        bool bMarked
        jointRx jJointRx = {j1=-132.269491, j2=127.123938, j3=-106.855674, j4=181.429188, j5=21.342688, j6=130.953129}
        pointRx pInter
        paraItem pParaItem
          [0]
            bool bSafePoint
            ifItem iIfItem
              [0]
                bool bANDOR[2]
                num nSigIndex[3]
                num nSigType[3]
                num nValue[3]
            mdesc mMdesc
            num nActionIndex = 42
            num nDelay
            num nMoveType = 1
            num nPercentage
            num nSigValue = 1
        pointRx pPointRx[2] = {x=-320.674662, y=-420.382638, z=642.0718966, rx=-1.140431, ry=0.333681, rz=-179.976981, shoulder=lefty, elbow=enegative, wrist=wpositive}
        string sID
      [45]
        bool bMarked
        jointRx jJointRx = {j1=-142.441106, j2=120.824327, j3=-88.705493, j4=181.282913, j5=33.0850501, j6=141.380041}
        pointRx pInter
        paraItem pParaItem
          [0]
            bool bSafePoint
            ifItem iIfItem
              [0]
                bool bANDOR[2]
                num nSigIndex[3]
                num nSigType[3]
                num nValue[3]
            mdesc mMdesc
            num nActionIndex = 42
            num nDelay
            num nMoveType = 1
            num nPercentage
            num nSigValue = 1
        pointRx pPointRx[2] = {x=-474.689621, y=-420.382631, z=642.0718894, rx=-1.140119, ry=0.333784, rz=-179.976923, shoulder=lefty, elbow=enegative, wrist=wpositive}
        string sID
      [46]
        bool bMarked
        jointRx jJointRx = {j1=-138.108258, j2=121.207146, j3=-89.710766, j4=181.162609, j5=32.51161, j6=137.142341}
        pointRx pInter
        paraItem pParaItem
          [0]
            bool bSafePoint
            ifItem iIfItem
              [0]
                bool bANDOR[2]
                num nSigIndex[3]
                num nSigType[3]
                num nValue[3]
            mdesc mMdesc
            num nActionIndex = 42
            num nDelay
            num nMoveType = 1
            num nPercentage
            num nSigValue = 1
        pointRx pPointRx[2] = {x=-436.796862, y=-451.644484, z=642.07189, rx=-1.139469, ry=0.334472, rz=-179.976638, shoulder=lefty, elbow=enegative, wrist=wpositive}
        string sID
      [47]
        bool bMarked
        jointRx jJointRx = {j1=-127.70596, j2=126.693595, j3=-105.454305, j4=181.135682, j5=22.350888, j6=126.671469}
        pointRx pInter
        paraItem pParaItem
          [0]
            bool bSafePoint
            ifItem iIfItem
              [0]
                bool bANDOR[2]
                num nSigIndex[3]
                num nSigType[3]
                num nValue[3]
            mdesc mMdesc
            num nActionIndex = 42
            num nDelay
            num nMoveType = 1
            num nPercentage
            num nSigValue = 1
        pointRx pPointRx[2] = {x=-290.683508, y=-451.609469, z=642.07191, rx=-1.140457, ry=0.335724, rz=-179.976594, shoulder=lefty, elbow=enegative, wrist=wpositive}
        string sID
      [48]
        bool bMarked
        jointRx jJointRx = {j1=-77.238254, j2=129.340507, j3=-114.913945, j4=177.831104, j5=15.475362, j6=79.35375}
        pointRx pInter
        paraItem pParaItem
          [0]
            bool bSafePoint
            ifItem iIfItem
              [0]
                bool bANDOR[2]
                num nSigIndex[3]
                num nSigType[3]
                num nValue[3]
            mdesc mMdesc
            num nActionIndex = 42
            num nDelay
            num nMoveType = 1
            num nPercentage
            num nSigValue = 1
        pointRx pPointRx[2] = {x=158.729452, y=-451.609464, z=642.0719065, rx=-1.140389, ry=0.334964, rz=-179.976748, shoulder=lefty, elbow=enegative, wrist=wpositive}
        string sID
      [49]
        bool bMarked
        jointRx jJointRx = {j1=-63.488687, j2=124.208026, j3=-97.940675, j4=178.228458, j5=27.14867, j6=65.0910716}
        pointRx pInter
        paraItem pParaItem
          [0]
            bool bSafePoint
            ifItem iIfItem
              [0]
                bool bANDOR[2]
                num nSigIndex[3]
                num nSigType[3]
                num nValue[3]
            mdesc mMdesc
            num nActionIndex = 42
            num nDelay
            num nMoveType = 1
            num nPercentage
            num nSigValue = 1
        pointRx pPointRx[2] = {x=310.830797, y=-495.30753, z=642.0718875, rx=-1.139453, ry=0.33486, rz=-179.976891, shoulder=lefty, elbow=enegative, wrist=wpositive}
        string sID
      [50]
        bool bMarked
        jointRx jJointRx = {j1=-78.0579912, j2=127.559769, j3=-108.316642, j4=178.378161, j5=20.297351, j6=79.604006}
        pointRx pInter
        paraItem pParaItem
          [0]
            bool bSafePoint
            ifItem iIfItem
              [0]
                bool bANDOR[2]
                num nSigIndex[3]
                num nSigType[3]
                num nValue[3]
            mdesc mMdesc
            num nActionIndex = 42
            num nDelay
            num nMoveType = 1
            num nPercentage
            num nSigValue = 1
        pointRx pPointRx[2] = {x=160.873249, y=-495.272541, z=642.0719096, rx=-1.140489, ry=0.333782, rz=-179.976981, shoulder=lefty, elbow=enegative, wrist=wpositive}
        string sID
      [51]
        bool bMarked
        jointRx jJointRx = {j1=-83.970136, j2=129.00855342, j3=-113.590578, j4=181.751291, j5=14.32041, j6=-96.622719}
        pointRx pInter
        paraItem pParaItem
          [0]
            bool bSafePoint
            ifItem iIfItem
              [0]
                bool bANDOR[2]
                num nSigIndex[3]
                num nSigType[3]
                num nValue[3]
            mdesc mMdesc
            num nActionIndex = 42
            num nDelay
            num nMoveType = 1
            num nPercentage
            num nSigValue = 1
        pointRx pPointRx[2] = {x=98.789636, y=-495.232609, z=642.0875542, rx=1.143362, ry=-0.31475, rz=1.103019, shoulder=lefty, elbow=enegative, wrist=wpositive}
        string sID
      [52]
        bool bMarked
        jointRx jJointRx = {j1=-101.251443, j2=129.329307, j3=-114.876217, j4=180.377122, j5=13.270505, j6=-78.0149862}
        pointRx pInter
        paraItem pParaItem
          [0]
            bool bSafePoint
            ifItem iIfItem
              [0]
                bool bANDOR[2]
                num nSigIndex[3]
                num nSigType[3]
                num nValue[3]
            mdesc mMdesc
            num nActionIndex = 42
            num nDelay
            num nMoveType = 1
            num nPercentage
            num nSigValue = 1
        pointRx pPointRx[2] = {x=-48.311282, y=-495.232554, z=642.0875543, rx=1.143247, ry=-0.315683, rz=1.102879, shoulder=lefty, elbow=enegative, wrist=wpositive}
        string sID
      [53]
        bool bMarked
        jointRx jJointRx = {j1=-117.974593, j2=127.746571, j3=-108.963712, j4=179.150072, j5=17.626951, j6=-60.118292}
        pointRx pInter
        paraItem pParaItem
          [0]
            bool bSafePoint
            ifItem iIfItem
              [0]
                bool bANDOR[2]
                num nSigIndex[3]
                num nSigType[3]
                num nValue[3]
            mdesc mMdesc
            num nActionIndex = 42
            num nDelay
            num nMoveType = 1
            num nPercentage
            num nSigValue = 1
        pointRx pPointRx[2] = {x=-203.879984, y=-495.232578, z=642.0875477, rx=1.143192, ry=-0.315734, rz=1.102838, shoulder=lefty, elbow=enegative, wrist=wpositive}
        string sID
      [54]
        bool bMarked
        jointRx jJointRx = {j1=-130.30363, j2=123.943868, j3=-97.190977, j4=178.849142, j5=25.681002, j6=-47.564193}
        pointRx pInter
        paraItem pParaItem
          [0]
            bool bSafePoint
            ifItem iIfItem
              [0]
                bool bANDOR[2]
                num nSigIndex[3]
                num nSigType[3]
                num nValue[3]
            mdesc mMdesc
            num nActionIndex = 42
            num nDelay
            num nMoveType = 1
            num nPercentage
            num nSigValue = 1
        pointRx pPointRx[2] = {x=-348.772288, y=-495.232559, z=642.0875407, rx=1.143488, ry=-0.315869, rz=1.102811, shoulder=lefty, elbow=enegative, wrist=wpositive}
        string sID
      [55]
        bool bMarked
        jointRx jJointRx = {j1=-87.553471, j2=145.12737, j3=-83.0900686, j4=182.117938, j5=63.691767, j6=-64.957345}
        pointRx pInter
        paraItem pParaItem
          [0]
            bool bSafePoint
            ifItem iIfItem
              [0]
                bool bANDOR[2]
                num nSigIndex[3]
                num nSigType[3]
                num nValue[3]
            mdesc mMdesc
            num nActionIndex = 42
            num nDelay
            num nMoveType = 1
            num nPercentage
            num nSigValue = 1
        pointRx pPointRx[2] = {x=61.326125, y=-652.062172, z=350.121525, rx=-1.556374, ry=-1.966704, rz=28.428639, shoulder=lefty, elbow=enegative, wrist=wpositive}
        string sID
    string sID
  [Position8_point_blow]
    num nFrameIndex
    num nMoveID
    num nToolIndex
    pointItem pPointItem[50]
      [0]
        bool bMarked
        jointRx jJointRx
        pointRx pInter
        paraItem pParaItem
          [0]
            bool bSafePoint
            ifItem iIfItem
              [0]
                bool bANDOR[2]
                num nSigIndex[3]
                num nSigType[3]
                num nValue[3]
            mdesc mMdesc
            num nActionIndex = 43
            num nDelay
            num nMoveType = 4
            num nPercentage
            num nSigValue = 1
        pointRx pPointRx[2]
        string sID
      [1]
        bool bMarked
        jointRx jJointRx = {j1=-87.553471, j2=145.12737, j3=-83.0900679, j4=182.117938, j5=63.691768, j6=-64.957345}
        pointRx pInter
        paraItem pParaItem
          [0]
            bool bSafePoint
            ifItem iIfItem
              [0]
                bool bANDOR[2]
                num nSigIndex[3]
                num nSigType[3]
                num nValue[3]
            mdesc mMdesc
            num nActionIndex = 42
            num nDelay
            num nMoveType = 1
            num nPercentage
            num nSigValue = 1
        pointRx pPointRx[2] = {x=61.326125, y=-652.062172, z=350.121525, rx=-1.556374, ry=-1.966704, rz=28.428639, shoulder=lefty, elbow=enegative, wrist=wpositive}
        string sID
      [2]
        bool bMarked
        jointRx jJointRx = {j1=-58.11069, j2=109.524278, j3=-71.857715, j4=179.347561, j5=40.141515, j6=-122.34843}
        pointRx pInter
        paraItem pParaItem
          [0]
            bool bSafePoint
            ifItem iIfItem
              [0]
                bool bANDOR[2]
                num nSigIndex[3]
                num nSigType[3]
                num nValue[3]
            mdesc mMdesc
            num nActionIndex = 42
            num nDelay
            num nMoveType = 1
            num nPercentage
            num nSigValue = 1
        pointRx pPointRx[2] = {x=409.39132, y=-556.393527, z=693.904783, rx=-2.322296, ry=-0.948981, rz=-0.986203, shoulder=lefty, elbow=enegative, wrist=wpositive}
        string sID
      [3]
        bool bMarked
        jointRx jJointRx = {j1=-66.225547, j2=113.999088, j3=-83.778734, j4=179.876465, j5=32.728091, j6=-114.636276}
        pointRx pInter
        paraItem pParaItem
          [0]
            bool bSafePoint
            ifItem iIfItem
              [0]
                bool bANDOR[2]
                num nSigIndex[3]
                num nSigType[3]
                num nValue[3]
            mdesc mMdesc
            num nActionIndex = 42
            num nDelay
            num nMoveType = 1
            num nPercentage
            num nSigValue = 1
        pointRx pPointRx[2] = {x=300.386557, y=-556.417777, z=693.904772, rx=-2.32202, ry=-0.949536, rz=-0.986453, shoulder=lefty, elbow=enegative, wrist=wpositive}
        string sID
      [4]
        bool bMarked
        jointRx jJointRx = {j1=-76.687433, j2=116.715992, j3=-91.802088, j4=180.847193, j5=27.394171, j6=-105.0405035}
        pointRx pInter
        paraItem pParaItem
          [0]
            bool bSafePoint
            ifItem iIfItem
              [0]
                bool bANDOR[2]
                num nSigIndex[3]
                num nSigType[3]
                num nValue[3]
            mdesc mMdesc
            num nActionIndex = 42
            num nDelay
            num nMoveType = 1
            num nPercentage
            num nSigValue = 1
        pointRx pPointRx[2] = {x=180.521932, y=-560.5436, z=693.904726, rx=-2.321521, ry=-0.949691, rz=-0.986547, shoulder=lefty, elbow=enegative, wrist=wpositive}
        string sID
      [5]
        bool bMarked
        jointRx jJointRx = {j1=-85.620281, j2=117.92465, j3=-95.696322, j4=181.846877, j5=24.627005, j6=-97.0419871}
        pointRx pInter
        paraItem pParaItem
          [0]
            bool bSafePoint
            ifItem iIfItem
              [0]
                bool bANDOR[2]
                num nSigIndex[3]
                num nSigType[3]
                num nValue[3]
            mdesc mMdesc
            num nActionIndex = 42
            num nDelay
            num nMoveType = 1
            num nPercentage
            num nSigValue = 1
        pointRx pPointRx[2] = {x=86.341042, y=-560.508796, z=693.904766, rx=-2.321719, ry=-0.949521, rz=-0.986489, shoulder=lefty, elbow=enegative, wrist=wpositive}
        string sID
      [6]
        bool bMarked
        jointRx jJointRx = {j1=-101.0757166, j2=116.15458, j3=-90.0727261, j4=182.913944, j5=28.207981, j6=-82.484873}
        pointRx pInter
        paraItem pParaItem
          [0]
            bool bSafePoint
            ifItem iIfItem
              [0]
                bool bANDOR[2]
                num nSigIndex[3]
                num nSigType[3]
                num nValue[3]
            mdesc mMdesc
            num nActionIndex = 42
            num nDelay
            num nMoveType = 1
            num nPercentage
            num nSigValue = 1
        pointRx pPointRx[2] = {x=-77.997367, y=-596.182081, z=693.904723, rx=-2.320616, ry=-0.948845, rz=-0.986256, shoulder=lefty, elbow=enegative, wrist=wpositive}
        string sID
      [7]
        bool bMarked
        jointRx jJointRx = {j1=-100.388707, j2=113.501769, j3=-82.38876, j4=182.465739, j5=33.248966, j6=-82.665703}
        pointRx pInter
        paraItem pParaItem
          [0]
            bool bSafePoint
            ifItem iIfItem
              [0]
                bool bANDOR[2]
                num nSigIndex[3]
                num nSigType[3]
                num nValue[3]
            mdesc mMdesc
            num nActionIndex = 42
            num nDelay
            num nMoveType = 1
            num nPercentage
            num nSigValue = 1
        pointRx pPointRx[2] = {x=-77.997368, y=-637.319122, z=693.904719, rx=-2.320623, ry=-0.948795, rz=-0.986246, shoulder=lefty, elbow=enegative, wrist=wpositive}
        string sID
      [8]
        bool bMarked
        jointRx jJointRx = {j1=-112.569059, j2=111.105712, j3=-75.937343, j4=182.939146, j5=36.983748, j6=-70.774258}
        pointRx pInter
        paraItem pParaItem
          [0]
            bool bSafePoint
            ifItem iIfItem
              [0]
                bool bANDOR[2]
                num nSigIndex[3]
                num nSigType[3]
                num nValue[3]
            mdesc mMdesc
            num nActionIndex = 42
            num nDelay
            num nMoveType = 1
            num nPercentage
            num nSigValue = 1
        pointRx pPointRx[2] = {x=-227.428005, y=-637.284544, z=693.904751, rx=-2.321115, ry=-0.949679, rz=-0.986554, shoulder=lefty, elbow=enegative, wrist=wpositive}
        string sID
      [9]
        bool bMarked
        jointRx jJointRx = {j1=-113.957376, j2=114.00103433, j3=-83.784205, j4=183.416468, j5=32.000017554, j6=-69.935449}
        pointRx pInter
        paraItem pParaItem
          [0]
            bool bSafePoint
            ifItem iIfItem
              [0]
                bool bANDOR[2]
                num nSigIndex[3]
                num nSigType[3]
                num nValue[3]
            mdesc mMdesc
            num nActionIndex = 42
            num nDelay
            num nMoveType = 1
            num nPercentage
            num nSigValue = 1
        pointRx pPointRx[2] = {x=-227.392618, y=-596.00613787, z=693.904773, rx=-2.322353, ry=-0.948517, rz=-0.986316, shoulder=lefty, elbow=enegative, wrist=wpositive}
        string sID
      [10]
        bool bMarked
        jointRx jJointRx = {j1=-131.107782, j2=122.205733, j3=-114.25278, j4=193.937243, j5=9.352415, j6=-63.640524}
        pointRx pInter
        paraItem pParaItem
          [0]
            bool bSafePoint
            ifItem iIfItem
              [0]
                bool bANDOR[2]
                num nSigIndex[3]
                num nSigType[3]
                num nValue[3]
            mdesc mMdesc
            num nActionIndex = 42
            num nDelay
            num nMoveType = 1
            num nPercentage
            num nSigValue = 1
        pointRx pPointRx[2] = {x=-278.571769, y=-365.527339, z=693.923849, rx=-2.325235, ry=-0.948268, rz=-0.986383, shoulder=lefty, elbow=enegative, wrist=wpositive}
        string sID
      [11]
        bool bMarked
        jointRx jJointRx = {j1=-135.395911, j2=104.707172, j3=-76.504799, j4=184.753699, j5=29.243911, j6=-49.740588}
        pointRx pInter
        paraItem pParaItem
          [0]
            bool bSafePoint
            ifItem iIfItem
              [0]
                bool bANDOR[2]
                num nSigIndex[3]
                num nSigType[3]
                num nValue[3]
            mdesc mMdesc
            num nActionIndex = 42
            num nDelay
            num nMoveType = 1
            num nPercentage
            num nSigValue = 1
        pointRx pPointRx[2] = {x=-444.435288, y=-480.130514, z=766.167371, rx=-2.324241, ry=-0.947818, rz=-0.986236, shoulder=lefty, elbow=enegative, wrist=wpositive}
        string sID
      [12]
        bool bMarked
        jointRx jJointRx = {j1=-134.796217, j2=92.950158, j3=-65.644872, j4=184.86577, j5=28.374058, j6=-50.474125}
        pointRx pInter
        paraItem pParaItem
          [0]
            bool bSafePoint
            ifItem iIfItem
              [0]
                bool bANDOR[2]
                num nSigIndex[3]
                num nSigType[3]
                num nValue[3]
            mdesc mMdesc
            num nActionIndex = 42
            num nDelay
            num nMoveType = 1
            num nPercentage
            num nSigValue = 1
        pointRx pPointRx[2] = {x=-444.435359, y=-489.966612, z=855.290958, rx=-2.324744, ry=-0.947384, rz=-0.986218, shoulder=lefty, elbow=enegative, wrist=wpositive}
        string sID
      [13]
        bool bMarked
        jointRx jJointRx = {j1=-136.173853, j2=87.871737, j3=-63.130701, j4=185.374273, j5=25.767564, j6=-49.65473}
        pointRx pInter
        paraItem pParaItem
          [0]
            bool bSafePoint
            ifItem iIfItem
              [0]
                bool bANDOR[2]
                num nSigIndex[3]
                num nSigType[3]
                num nValue[3]
            mdesc mMdesc
            num nActionIndex = 42
            num nDelay
            num nMoveType = 1
            num nPercentage
            num nSigValue = 1
        pointRx pPointRx[2] = {x=-444.435358, y=-467.674325, z=901.291627, rx=-2.325949, ry=-0.946701, rz=-0.986341, shoulder=lefty, elbow=enegative, wrist=wpositive}
        string sID
      [14]
        bool bMarked
        jointRx jJointRx = {j1=-141.164951, j2=86.59666, j3=-69.357957, j4=187.756915, j5=18.114888, j6=-47.194082}
        pointRx pInter
        paraItem pParaItem
          [0]
            bool bSafePoint
            ifItem iIfItem
              [0]
                bool bANDOR[2]
                num nSigIndex[3]
                num nSigType[3]
                num nValue[3]
            mdesc mMdesc
            num nActionIndex = 42
            num nDelay
            num nMoveType = 1
            num nPercentage
            num nSigValue = 1
        pointRx pPointRx[2] = {x=-444.435342, y=-395.0345733, z=930.658223, rx=-2.325698, ry=-0.946616, rz=-0.986323, shoulder=lefty, elbow=enegative, wrist=wpositive}
        string sID
      [15]
        bool bMarked
        jointRx jJointRx = {j1=-150.996048, j2=88.749744, j3=-81.786263, j4=199.00922873, j5=7.675391, j6=-48.828489}
        pointRx pInter
        paraItem pParaItem
          [0]
            bool bSafePoint
            ifItem iIfItem
              [0]
                bool bANDOR[2]
                num nSigIndex[3]
                num nSigType[3]
                num nValue[3]
            mdesc mMdesc
            num nActionIndex = 42
            num nDelay
            num nMoveType = 1
            num nPercentage
            num nSigValue = 1
        pointRx pPointRx[2] = {x=-444.435068, y=-278.693508, z=930.65815, rx=-2.325239, ry=-0.948289, rz=-0.986304, shoulder=lefty, elbow=enegative, wrist=wpositive}
        string sID
      [16]
        bool bMarked
        jointRx jJointRx = {j1=-136.944318, j2=108.102124, j3=-81.594441, j4=185.0858237, j5=27.496189, j6=-48.554881}
        pointRx pInter
        paraItem pParaItem
          [0]
            bool bSafePoint
            ifItem iIfItem
              [0]
                bool bANDOR[2]
                num nSigIndex[3]
                num nSigType[3]
                num nValue[3]
            mdesc mMdesc
            num nActionIndex = 42
            num nDelay
            num nMoveType = 1
            num nPercentage
            num nSigValue = 1
        pointRx pPointRx[2] = {x=-444.435337, y=-455.673073, z=747.789181, rx=-2.325621, ry=-0.946829, rz=-0.986212, shoulder=lefty, elbow=enegative, wrist=wpositive}
        string sID
      [17]
        bool bMarked
        jointRx jJointRx = {j1=-133.102266, j2=114.394979, j3=-110.124586, j4=185.156231, j5=6.735085, j6=-104.330607}
        pointRx pInter
        paraItem pParaItem
          [0]
            bool bSafePoint
            ifItem iIfItem
              [0]
                bool bANDOR[2]
                num nSigIndex[3]
                num nSigType[3]
                num nValue[3]
            mdesc mMdesc
            num nActionIndex = 42
            num nDelay
            num nMoveType = 1
            num nPercentage
            num nSigValue = 1
        pointRx pPointRx[2] = {x=-273.0764108, y=-357.254112, z=747.804416, rx=-2.192889, ry=1.224247, rz=-52.275755, shoulder=lefty, elbow=enegative, wrist=wpositive}
        string sID
      [18]
        bool bMarked
        jointRx jJointRx = {j1=-117.270513, j2=113.78497, j3=-104.717978, j4=179.481532, j5=11.577034, j6=-114.962229}
        pointRx pInter
        paraItem pParaItem
          [0]
            bool bSafePoint
            ifItem iIfItem
              [0]
                bool bANDOR[2]
                num nSigIndex[3]
                num nSigType[3]
                num nValue[3]
            mdesc mMdesc
            num nActionIndex = 42
            num nDelay
            num nMoveType = 1
            num nPercentage
            num nSigValue = 1
        pointRx pPointRx[2] = {x=-176.508441, y=-453.51729, z=747.804419, rx=-2.183299, ry=1.242081, rz=-52.719273, shoulder=lefty, elbow=enegative, wrist=wpositive}
        string sID
      [19]
        bool bMarked
        jointRx jJointRx = {j1=-109.137554, j2=109.619736, j3=-86.542307, j4=178.941557, j5=25.551631, j6=-122.640865}
        pointRx pInter
        paraItem pParaItem
          [0]
            bool bSafePoint
            ifItem iIfItem
              [0]
                bool bANDOR[2]
                num nSigIndex[3]
                num nSigType[3]
                num nValue[3]
            mdesc mMdesc
            num nActionIndex = 42
            num nDelay
            num nMoveType = 1
            num nPercentage
            num nSigValue = 1
        pointRx pPointRx[2] = {x=-144.182021, y=-580.158289, z=747.804426, rx=-2.184454, ry=1.240986, rz=-52.719545, shoulder=lefty, elbow=enegative, wrist=wpositive}
        string sID
      [20]
        bool bMarked
        jointRx jJointRx = {j1=-105.96936, j2=113.946894, j3=-105.873919, j4=176.762051, j5=10.531462, j6=-123.577788}
        pointRx pInter
        paraItem pParaItem
          [0]
            bool bSafePoint
            ifItem iIfItem
              [0]
                bool bANDOR[2]
                num nSigIndex[3]
                num nSigType[3]
                num nValue[3]
            mdesc mMdesc
            num nActionIndex = 42
            num nDelay
            num nMoveType = 1
            num nPercentage
            num nSigValue = 1
        pointRx pPointRx[2] = {x=-78.145175, y=-473.574291, z=747.804414, rx=-2.185277, ry=1.240398, rz=-52.719616, shoulder=lefty, elbow=enegative, wrist=wpositive}
        string sID
      [21]
        bool bMarked
        jointRx jJointRx = {j1=-100.135452, j2=114.341428, j3=-109.460145, j4=173.401757, j5=7.298155, j6=-126.0452472}
        pointRx pInter
        paraItem pParaItem
          [0]
            bool bSafePoint
            ifItem iIfItem
              [0]
                bool bANDOR[2]
                num nSigIndex[3]
                num nSigType[3]
                num nValue[3]
            mdesc mMdesc
            num nActionIndex = 42
            num nDelay
            num nMoveType = 1
            num nPercentage
            num nSigValue = 1
        pointRx pPointRx[2] = {x=-23.263146, y=-455.736187, z=747.804388, rx=-2.18503, ry=1.240118, rz=-52.719596, shoulder=lefty, elbow=enegative, wrist=wpositive}
        string sID
      [22]
        bool bMarked
        jointRx jJointRx = {j1=-100.135452, j2=114.341428, j3=-109.460145, j4=173.401757, j5=7.298155, j6=-126.0452472}
        pointRx pInter
        paraItem pParaItem
          [0]
            bool bSafePoint
            ifItem iIfItem
              [0]
                bool bANDOR[2]
                num nSigIndex[3]
                num nSigType[3]
                num nValue[3]
            mdesc mMdesc
            num nActionIndex = 42
            num nDelay
            num nMoveType
            num nPercentage
            num nSigValue = 1
        pointRx pPointRx[2] = {x=-23.263146, y=-455.736187, z=747.804388, rx=-2.18503, ry=1.240118, rz=-52.719596, shoulder=lefty, elbow=enegative, wrist=wpositive}
        string sID
      [23]
        bool bMarked
        jointRx jJointRx = {j1=-106.631553, j2=109.786963, j3=-134.970625, j4=184.819916, j5=-24.691551, j6=-80.199638}
        pointRx pInter
        paraItem pParaItem
          [0]
            bool bSafePoint
            ifItem iIfItem
              [0]
                bool bANDOR[2]
                num nSigIndex[3]
                num nSigType[3]
                num nValue[3]
            mdesc mMdesc
            num nActionIndex = 42
            num nDelay
            num nMoveType
            num nPercentage
            num nSigValue = 1
        pointRx pPointRx[2] = {x=-10.865105, y=-272.383063, z=740.397718, rx=0.0307126, ry=2.090166, rz=-2.46071, shoulder=lefty, elbow=enegative, wrist=wnegative}
        string sID
      [24]
        bool bMarked
        jointRx jJointRx = {j1=-81.325877, j2=110.844378, j3=-133.586221, j4=185.246198, j5=-23.174992, j6=-105.96506}
        pointRx pInter
        paraItem pParaItem
          [0]
            bool bSafePoint
            ifItem iIfItem
              [0]
                bool bANDOR[2]
                num nSigIndex[3]
                num nSigType[3]
                num nValue[3]
            mdesc mMdesc
            num nActionIndex = 42
            num nDelay
            num nMoveType = 1
            num nPercentage
            num nSigValue = 1
        pointRx pPointRx[2] = {x=110.33304, y=-272.382932, z=740.397731, rx=0.0311611, ry=2.0907781, rz=-2.460321, shoulder=lefty, elbow=enegative, wrist=wnegative}
        string sID
      [25]
        bool bMarked
        jointRx jJointRx = {j1=-96.0712223, j2=114.244351, j3=-126.542039, j4=186.250879, j5=-10.611959, j6=-41.0712755}
        pointRx pInter
        paraItem pParaItem
          [0]
            bool bSafePoint
            ifItem iIfItem
              [0]
                bool bANDOR[2]
                num nSigIndex[3]
                num nSigType[3]
                num nValue[3]
            mdesc mMdesc
            num nActionIndex = 42
            num nDelay
            num nMoveType = 1
            num nPercentage
            num nSigValue = 1
        pointRx pPointRx[2] = {x=24.601437, y=-336.239263, z=740.397725, rx=-1.61612, ry=1.32728, rz=49.00349569, shoulder=lefty, elbow=enegative, wrist=wnegative}
        string sID
      [26]
        bool bMarked
        jointRx jJointRx = {j1=-95.690534, j2=114.696488, j3=-124.883411, j4=183.926416, j5=-8.191559, j6=-21.0119831}
        pointRx pInter
        paraItem pParaItem
          [0]
            bool bSafePoint
            ifItem iIfItem
              [0]
                bool bANDOR[2]
                num nSigIndex[3]
                num nSigType[3]
                num nValue[3]
            mdesc mMdesc
            num nActionIndex = 42
            num nDelay
            num nMoveType = 1
            num nPercentage
            num nSigValue = 1
        pointRx pPointRx[2] = {x=20.559143, y=-347.136674, z=740.39771, rx=-1.949012, ry=0.755958, rz=67.186994, shoulder=lefty, elbow=enegative, wrist=wnegative}
        string sID
      [27]
        bool bMarked
        jointRx jJointRx = {j1=-100.882638, j2=115.524729, j3=-119.715858, j4=189.99726, j5=-2.166253, j6=-21.927142}
        pointRx pInter
        paraItem pParaItem
          [0]
            bool bSafePoint
            ifItem iIfItem
              [0]
                bool bANDOR[2]
                num nSigIndex[3]
                num nSigType[3]
                num nValue[3]
            mdesc mMdesc
            num nActionIndex = 42
            num nDelay
            num nMoveType = 1
            num nPercentage
            num nSigValue = 1
        pointRx pPointRx[2] = {x=-20.271174, y=-387.650591, z=740.397525, rx=-1.949817, ry=0.75764, rz=67.18662, shoulder=lefty, elbow=enegative, wrist=wnegative}
        string sID
      [28]
        bool bMarked
        jointRx jJointRx = {j1=-98.590862, j2=115.394944, j3=-120.62517, j4=152.249394, j5=-3.377524, j6=83.0398225}
        pointRx pInter
        paraItem pParaItem
          [0]
            bool bSafePoint
            ifItem iIfItem
              [0]
                bool bANDOR[2]
                num nSigIndex[3]
                num nSigType[3]
                num nValue[3]
            mdesc mMdesc
            num nActionIndex = 42
            num nDelay
            num nMoveType = 1
            num nPercentage
            num nSigValue = 1
        pointRx pPointRx[2] = {x=-20.237233, y=-376.857663, z=740.396708, rx=-2.449976, ry=-1.219744, rz=136.744035, shoulder=lefty, elbow=enegative, wrist=wnegative}
        string sID
      [29]
        bool bMarked
        jointRx jJointRx = {j1=-94.342198, j2=115.399464, j3=-120.574953, j4=153.574077, j5=-3.150419, j6=77.473821}
        pointRx pInter
        paraItem pParaItem
          [0]
            bool bSafePoint
            ifItem iIfItem
              [0]
                bool bANDOR[2]
                num nSigIndex[3]
                num nSigType[3]
                num nValue[3]
            mdesc mMdesc
            num nActionIndex = 42
            num nDelay
            num nMoveType = 1
            num nPercentage
            num nSigValue = 1
        pointRx pPointRx[2] = {x=9.265961, y=-376.836715, z=740.402193, rx=-2.45298, ry=-1.219325, rz=136.742906, shoulder=lefty, elbow=enegative, wrist=wnegative}
        string sID
      [30]
        bool bMarked
        jointRx jJointRx = {j1=-98.415545, j2=115.64334, j3=-116.881458, j4=131.21052, j5=-3.390587, j6=180.414513}
        pointRx pInter
        paraItem pParaItem
          [0]
            bool bSafePoint
            ifItem iIfItem
              [0]
                bool bANDOR[2]
                num nSigIndex[3]
                num nSigType[3]
                num nValue[3]
            mdesc mMdesc
            num nActionIndex = 42
            num nDelay
            num nMoveType = 1
            num nPercentage
            num nSigValue = 1
        pointRx pPointRx[2] = {x=-35.863926, y=-432.0528257, z=740.403674, rx=0.613001, ry=-2.668531, rz=-146.748671, shoulder=lefty, elbow=enegative, wrist=wnegative}
        string sID
      [31]
        bool bMarked
        jointRx jJointRx = {j1=-101.750183, j2=114.53034, j3=-125.268384, j4=164.764824, j5=-9.193065, j6=150.0786226}
        pointRx pInter
        paraItem pParaItem
          [0]
            bool bSafePoint
            ifItem iIfItem
              [0]
                bool bANDOR[2]
                num nSigIndex[3]
                num nSigType[3]
                num nValue[3]
            mdesc mMdesc
            num nActionIndex = 42
            num nDelay
            num nMoveType = 1
            num nPercentage
            num nSigValue = 1
        pointRx pPointRx[2] = {x=-41.0858853, y=-339.972742, z=740.403727, rx=-2.313723, ry=-1.976447, rz=-146.720771, shoulder=lefty, elbow=enegative, wrist=wnegative}
        string sID
      [32]
        bool bMarked
        jointRx jJointRx = {j1=-93.176498, j2=114.397129, j3=-125.767117, j4=167.0222508, j5=-9.404252, j6=139.264507}
        pointRx pInter
        paraItem pParaItem
          [0]
            bool bSafePoint
            ifItem iIfItem
              [0]
                bool bANDOR[2]
                num nSigIndex[3]
                num nSigType[3]
                num nValue[3]
            mdesc mMdesc
            num nActionIndex = 42
            num nDelay
            num nMoveType = 1
            num nPercentage
            num nSigValue = 1
        pointRx pPointRx[2] = {x=13.0926046, y=-335.307093, z=740.403563, rx=-2.31492, ry=-1.977735, rz=-146.720656, shoulder=lefty, elbow=enegative, wrist=wnegative}
        string sID
      [33]
        bool bMarked
        jointRx jJointRx = {j1=-92.339418, j2=114.605155, j3=-124.971473, j4=176.0737376, j5=-7.38225, j6=96.22607}
        pointRx pInter
        paraItem pParaItem
          [0]
            bool bSafePoint
            ifItem iIfItem
              [0]
                bool bANDOR[2]
                num nSigIndex[3]
                num nSigType[3]
                num nValue[3]
            mdesc mMdesc
            num nActionIndex = 42
            num nDelay
